(*!
<summary>Reports the outcome of copying a mapped source into existing generic value storage.</summary>
*)
(*
SPDX-FileCopyrightText: © 2026 Oleksandr Tiutyk <trofimich@gmail.com>
SPDX-License-Identifier: MIT
License: https://opensource.org/license/mit
*)

{attribute 'qualified_only'}
{attribute 'strict'}
{attribute 'to_string'}
TYPE GENERIC_VALUE_COPY_RESULT :
(
	COPIED,
	INCOMPATIBLE_TYPE,
	INSUFFICIENT_CAPACITY,
	COPY_FAILED
);
END_TYPE

(* stored: Version 1.1.0.1
   DUT GENERIC_VALUE_COPY_RESULT: Id {35ea289b-5678-41e4-a703-b8100f4f73f1} *)
